(*
SPDX-FileCopyrightText: © 2026 Oleksandr Tiutyk <trofimich@gmail.com>
SPDX-License-Identifier: MIT
License: https://opensource.org/license/mit
*)

(*!
<summary>Holds one pending operand check during a synchronous workflow load.</summary>
<description>The loader owns the entry and borrows its scope until validation or rollback.</description>
*)

{attribute 'enable_dynamic_creation'}		
TYPE VARIABLE_REQUIREMENT :
STRUCT
	Scope : IVariableLookup;
	Name : STRING;
	Next : POINTER TO VARIABLE_REQUIREMENT;
END_STRUCT
END_TYPE

(* stored: Version 1.1.0.1
   DUT VARIABLE_REQUIREMENT: Id {55ca11f3-e8f1-48d9-8dcc-a2a65975a8b7} *)
